(* IEC 61131-3 sources: rusty/tests/lit/single/string_functions, 5 files *)

(* ---- concat.st ---- *)
// RUN: %COMPILE %s && %RUN | %CHECK %s
// End-to-end tests for the CONCAT stdlib function (STRING and WSTRING).
// Also covers truncation to the STRING[2048] / WSTRING[2048] result buffer:
// concatenating past 2048 code units used to overflow the result buffer and
// crash; it must now truncate to 2048 instead. See libs/stdlib/src/string_functions.rs.

FUNCTION main : DINT
VAR
    s      : STRING[2048];
    ws     : WSTRING[2048];
    chunk  : STRING[2048]  := 'AAAAAAAAAAAAAAAAAAAAAAAAAAAAAAAAAAAAAAAAAAAAAAAAAAAAAAAAAAAAAAAAAAAAAAAAAAAAAAAAAAAAAAAAAAAAAAAAAAAAAAAAAAAAAAAAAAAAAAAAAAAAAAAA';
    wchunk : WSTRING[2048] := "AAAAAAAAAAAAAAAAAAAAAAAAAAAAAAAAAAAAAAAAAAAAAAAAAAAAAAAAAAAAAAAAAAAAAAAAAAAAAAAAAAAAAAAAAAAAAAAAAAAAAAAAAAAAAAAAAAAAAAAAAAAAAAAA";
    big    : STRING[2048];
    wbig   : WSTRING[2048];
END_VAR
    // --- functional: STRING ---
    s := CONCAT('Hello', ', ', 'World', '!');
    // CHECK: Hello, World!
    printf('%s$N', REF(s));

    // --- functional: WSTRING ---
    ws := CONCAT("Hello", ", ", "World", "!");
    // CHECK: Hello, World!
    printf('%s$N', REF(TO_STRING(ws)));

    // --- truncation: STRING ---
    // 16 * 128 == 2048 fills the buffer exactly (no truncation yet).
    big := CONCAT(chunk, chunk, chunk, chunk, chunk, chunk, chunk, chunk, chunk, chunk, chunk, chunk, chunk, chunk, chunk, chunk);
    // CHECK: 2048
    printf('%d$N', LEN(big));
    // CONCAT(big, big) would be 4096; must truncate to 2048 instead of crashing.
    s := CONCAT(big, big);
    // CHECK: 2048
    printf('%d$N', LEN(s));

    // --- truncation: WSTRING ---
    wbig := CONCAT(wchunk, wchunk, wchunk, wchunk, wchunk, wchunk, wchunk, wchunk, wchunk, wchunk, wchunk, wchunk, wchunk, wchunk, wchunk, wchunk);
    ws := CONCAT(wbig, wbig);
    // CHECK: 2048
    printf('%d$N', LEN(ws));

    main := 0;
END_FUNCTION

(* ---- concat_scalar_generic_no_duplicate.st ---- *)
// RUN: not %COMPILE %s --error-format clang 2>&1 | %CHECK %s
// Regression: a nature violation on a generic function with a *scalar* return (here CONCAT_LTOD,
// `<T: ANY_INT> : LTOD`) must be reported exactly once. Such calls are NOT rewritten by the
// aggregate-return lowerer, so their generic nature survives to the regular validation pass. The
// lowerer must therefore stay silent for them; otherwise the diagnostic is emitted twice (once by
// the lowerer, once by validation). The CHECK-NEXT below pins the abort line directly after the
// single E062, so a duplicate E062 would fail the test.

FUNCTION mainProg : LTOD
VAR
    r : REAL;
    i : INT;
END_VAR
    // CHECK: {{.*}}error[E062]: Invalid type nature for generic argument. REAL is no ANY_INT
    // CHECK-NEXT: error: Compilation aborted due to critical errors
    mainProg := CONCAT_LTOD(r, i, i, i);
END_FUNCTION

(* ---- concat_type_mismatch.st ---- *)
// RUN: not %COMPILE %s --error-format clang 2>&1 | %CHECK %s
// End-to-end guard for passing non-string arguments to the generic CONCAT stdlib function.
// CONCAT is `FUNCTION CONCAT <T: ANY_STRING> : T` with a `{ref} {sized} T...` variadic. Passing a
// non-ANY_STRING argument used to compile silently and then crash in codegen: the generic call is
// lowered to the concrete `CONCAT__STRING` and the following re-annotation dropped the generic
// nature before validation could see it. Every offending argument must now be reported, while
// genuine string arguments are left alone.

FUNCTION mainProg : DINT
VAR
    x : DINT;
    y : REAL;
    z : STRING;
END_VAR
    // Every non-string argument is flagged individually; `z` is a valid STRING and is not.
    // CHECK-DAG: {{.*}}concat_type_mismatch.st:[[@LINE+1]]:{{[0-9]+}}:{{.*}}error[E062]: Invalid type nature for generic argument. DINT is no ANY_STRING
    z := CONCAT(x, z);

    // CHECK-DAG: {{.*}}concat_type_mismatch.st:[[@LINE+2]]:{{[0-9]+}}:{{.*}}error[E062]: Invalid type nature for generic argument. DINT is no ANY_STRING
    // CHECK-DAG: {{.*}}concat_type_mismatch.st:[[@LINE+1]]:{{[0-9]+}}:{{.*}}error[E062]: Invalid type nature for generic argument. REAL is no ANY_STRING
    z := CONCAT(x, y, z);
END_FUNCTION

(* ---- insert.st ---- *)
// RUN: %COMPILE %s && %RUN | %CHECK %s
// End-to-end tests for the INSERT stdlib function (STRING and WSTRING).
// INSERT combines two strings, so its result can exceed the STRING[2048] /
// WSTRING[2048] result buffer. That used to overflow the buffer and crash;
// it must now truncate to 2048 instead. See libs/stdlib/src/string_functions.rs.

FUNCTION main : DINT
VAR
    s      : STRING[2048];
    ws     : WSTRING[2048];
    chunk  : STRING[2048]  := 'AAAAAAAAAAAAAAAAAAAAAAAAAAAAAAAAAAAAAAAAAAAAAAAAAAAAAAAAAAAAAAAAAAAAAAAAAAAAAAAAAAAAAAAAAAAAAAAAAAAAAAAAAAAAAAAAAAAAAAAAAAAAAAAA';
    wchunk : WSTRING[2048] := "AAAAAAAAAAAAAAAAAAAAAAAAAAAAAAAAAAAAAAAAAAAAAAAAAAAAAAAAAAAAAAAAAAAAAAAAAAAAAAAAAAAAAAAAAAAAAAAAAAAAAAAAAAAAAAAAAAAAAAAAAAAAAAAA";
    big    : STRING[2048];
    wbig   : WSTRING[2048];
END_VAR
    // --- functional: STRING --- (keep the first 2 characters, then insert)
    s := INSERT('Hello', 'XYZ', 2);
    // CHECK: HeXYZllo
    printf('%s$N', REF(s));

    // --- functional: WSTRING ---
    ws := INSERT("Hello", "XYZ", 2);
    // CHECK: HeXYZllo
    printf('%s$N', REF(TO_STRING(ws)));

    // --- truncation: STRING ---
    big := CONCAT(chunk, chunk, chunk, chunk, chunk, chunk, chunk, chunk, chunk, chunk, chunk, chunk, chunk, chunk, chunk, chunk);
    // INSERT(big, big, 10) would be ~4096; must truncate to 2048.
    s := INSERT(big, big, 10);
    // CHECK: 2048
    printf('%d$N', LEN(s));

    // --- truncation: WSTRING ---
    wbig := CONCAT(wchunk, wchunk, wchunk, wchunk, wchunk, wchunk, wchunk, wchunk, wchunk, wchunk, wchunk, wchunk, wchunk, wchunk, wchunk, wchunk);
    ws := INSERT(wbig, wbig, 10);
    // CHECK: 2048
    printf('%d$N', LEN(ws));

    main := 0;
END_FUNCTION

(* ---- replace.st ---- *)
// RUN: %COMPILE %s && %RUN | %CHECK %s
// End-to-end tests for the REPLACE stdlib function (STRING and WSTRING).
// REPLACE can grow a string when the replacement is longer than the replaced
// region, so its result can exceed the STRING[2048] / WSTRING[2048] result
// buffer. That used to overflow the buffer and crash; it must now truncate to
// 2048 instead. See libs/stdlib/src/string_functions.rs.

FUNCTION main : DINT
VAR
    s      : STRING[2048];
    ws     : WSTRING[2048];
    chunk  : STRING[2048]  := 'AAAAAAAAAAAAAAAAAAAAAAAAAAAAAAAAAAAAAAAAAAAAAAAAAAAAAAAAAAAAAAAAAAAAAAAAAAAAAAAAAAAAAAAAAAAAAAAAAAAAAAAAAAAAAAAAAAAAAAAAAAAAAAAA';
    wchunk : WSTRING[2048] := "AAAAAAAAAAAAAAAAAAAAAAAAAAAAAAAAAAAAAAAAAAAAAAAAAAAAAAAAAAAAAAAAAAAAAAAAAAAAAAAAAAAAAAAAAAAAAAAAAAAAAAAAAAAAAAAAAAAAAAAAAAAAAAAA";
    big    : STRING[2048];
    wbig   : WSTRING[2048];
END_VAR
    // --- functional: STRING --- (replace 2 characters starting at position 2)
    s := REPLACE('Hello', 'XX', 2, 2);
    // CHECK: HXXlo
    printf('%s$N', REF(s));

    // --- functional: WSTRING ---
    ws := REPLACE("Hello", "XX", 2, 2);
    // CHECK: HXXlo
    printf('%s$N', REF(TO_STRING(ws)));

    // --- truncation: STRING ---
    big := CONCAT(chunk, chunk, chunk, chunk, chunk, chunk, chunk, chunk, chunk, chunk, chunk, chunk, chunk, chunk, chunk, chunk);
    // REPLACE(big, big, 1, 1) would be ~4095; must truncate to 2048.
    s := REPLACE(big, big, 1, 1);
    // CHECK: 2048
    printf('%d$N', LEN(s));

    // --- truncation: WSTRING ---
    wbig := CONCAT(wchunk, wchunk, wchunk, wchunk, wchunk, wchunk, wchunk, wchunk, wchunk, wchunk, wchunk, wchunk, wchunk, wchunk, wchunk, wchunk);
    ws := REPLACE(wbig, wbig, 1, 1);
    // CHECK: 2048
    printf('%d$N', LEN(ws));

    main := 0;
END_FUNCTION
